Yaskawa INFORM job: DEMO_RJ_XYZ.JBI

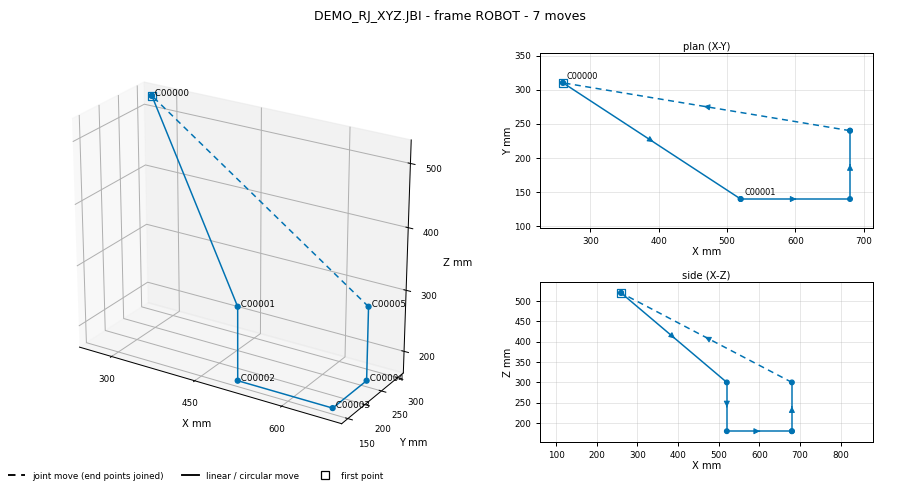
[picture p0: tool path of DEMO_RJ_XYZ.JBI in frame ROBOT, 7 of 7 moves have a stored position in this frame; points joined in program order, loops and branches not executed]
/JOB
//NAME DEMO_RJ_XYZ
//POS
///NPOS 7,0,0,0,0,0
///TOOL 8
///POSTYPE ROBOT
///RECTAN
///RCONF 0,0,1,0,0,0,0,0,0,0,0,0,0,0,0,0,0,0,0,0,0,0,0,0
C00000=260.000,310.000,520.000,-179.5000,1.2500,-12.0000
C00001=520.000,140.000,300.000,-179.5000,1.2500,25.0000
C00002=520.000,140.000,180.000,-179.5000,1.2500,25.0000
C00003=680.000,140.000,180.000,-179.5000,1.2500,25.0000
C00004=680.000,240.000,180.000,-179.5000,1.2500,25.0000
C00005=680.000,240.000,300.000,-179.5000,1.2500,25.0000
C00006=260.000,310.000,520.000,-179.5000,1.2500,-12.0000
//INST
///DATE 2026/11/03 16:00
///ATTR SC,RW,RJ
////FRAME ROBOT
///GROUP1 RB1
NOP
'SYNTHETIC DEMO JOB - NOT A REAL ROBOT JOB
MOVJ C00000 VJ=25.00
MOVL C00001 V=150.0
MOVL C00002 V=60.0
MOVL C00003 V=60.0
MOVL C00004 V=60.0
MOVL C00005 V=150.0
MOVJ C00006 VJ=25.00
END
